(* IEC 61131-3 sources: rusty/tests/lit/multi/build_info_dedup, 2 files *)

(* ---- helper.st ---- *)
FUNCTION standalone_helper : DINT
    standalone_helper := 42;
END_FUNCTION

(* ---- main.st ---- *)
FUNCTION main : DINT
    main := 0;
END_FUNCTION
